// CRONOMETRO: misura il tempo trascorso dall'ultimo Reset e lo confronta con una durata.
// Non serve chiamare il corpo del blocco: si usano solo metodi e action.
FUNCTION_BLOCK FB_Timer
VAR_INPUT
	tTimer		:	TIME;	// durata usata da VerifySelfElapsed
END_VAR
VAR
	tStartTime	:	TIME	:=	TIME() - tTimer;	// istante dell'ultimo Reset
END_VAR

// IMPOSTA LA DURATA USATA DA VerifySelfElapsed (non fa ripartire il cronometro)
METHOD ChangeTimer
VAR_INPUT
	tTimerNew	:	TIME;
END_VAR
tTimer	:=	tTimerNew;
END_METHOD

// TEMPO TRASCORSO DALL'ULTIMO RESET
METHOD ComputeElapsed : TIME
ComputeElapsed	:=	TIME() - tStartTime;
END_METHOD

// TEMPO TRASCORSO DALL'ULTIMO RESET, IN SECONDI
METHOD ComputeElapsedSeconds : REAL
VAR_INPUT
END_VAR
ComputeElapsedSeconds	:=	F_TimeToSeconds(ComputeElapsed());
END_METHOD

ACTION Reset:
// FA RIPARTIRE IL CRONOMETRO DA ZERO
tStartTime	:=	TIME();
END_ACTION

// FA RIPARTIRE IL CRONOMETRO SOLO SE bCondition È TRUE.
// Restituisce TRUE se il reset è stato eseguito.
METHOD ResetCondition : BOOL
VAR_INPUT
	bCondition	:	BOOL;
END_VAR
IF bCondition THEN
	Reset();
END_IF
ResetCondition	:=	bCondition;
END_METHOD

// FA RIPARTIRE IL CRONOMETRO COME SE FOSSE GIÀ TRASCORSO tOffset
METHOD ResetWithOffset
VAR_INPUT
	tOffset	:	TIME;
END_VAR
tStartTime	:=	TIME() - tOffset;
END_METHOD

// TRUE SE DALL'ULTIMO RESET È TRASCORSO PIÙ DI tInputTime
METHOD VerifyElapsed : BOOL
VAR_INPUT
	tInputTime	:	TIME;
END_VAR
VerifyElapsed	:=	ComputeElapsed() > tInputTime;
END_METHOD

// TRUE SE DALL'ULTIMO RESET È TRASCORSO PIÙ DI tTimer
METHOD VerifySelfElapsed : BOOL
VerifySelfElapsed	:=	ComputeElapsed() > tTimer;
END_METHOD

END_FUNCTION_BLOCK

(* stored: Version 1.1.0.1, ProductVersion 3.1.4024.9
   POU FB_Timer: Id {1c7e49d7-0b84-41e9-bf71-580086c34571}, SpecialFunc None
   Folder ACTIONs: Id {65ec57ae-aace-4f74-9168-933038335526}
   Folder METHODs: Id {b8755bcd-b80c-49c5-87a5-dae8f18a163c}
   Method ChangeTimer: Id {ec14ba12-8668-4679-91c7-1c207881d044}
   Method ComputeElapsed: Id {a50a418d-2f72-4912-800d-1c6a8b325b98}
   Method ComputeElapsedSeconds: Id {dbb68b9c-c223-4ea3-93c9-0ff1dcc37603}
   Action Reset: Id {82e45bc8-9b92-44a8-ae3c-9f0229c7d221}
   Method ResetCondition: Id {22784363-67a0-4843-8592-80fdd94ad69e}
   Method ResetWithOffset: Id {a9a5c184-95ea-4593-920b-fbd3201fa968}
   Method VerifyElapsed: Id {c27fb815-8bc4-4f79-9061-f28220489b90}
   Method VerifySelfElapsed: Id {8a8f8a9b-1b74-447b-aa6b-e346929972fb} *)
